SUBAPPLICATION SERVER_0_QO (* OPC-UA-Methode ohne Argumente (CREATE_METHOD): IND nur bei echtem Aufruf (QO=TRUE), RSP intern *)
  (* Standard: 61499-2; Description: Copyright (c) 2026 Meisterschulen am Ostbahnhof This program and the accompanying materials are made available under the terms of the Eclipse Public License 2.0 which is available at https://www.eclipse.org/legal/epl-2.0/ SPDX-License-Identifier: EPL-2.0 *)
  (* Version 1.0, 2026-11-25, Franz Höpfinger, Meisterschulen am Ostbahnhof, Neu: SERVER_0 + E_PERMIT(PERMIT=QO). Ein gescheitertes RSP meldet IND mit QO=FALSE, direkt IND->RSP ergab eine Endlosschleife. *)
  PACKAGE MyLib::net;
  (* Documentation:
  OPC-UA-Methode ohne Argumente, sicher beantwortet
   SERVER_0 mit CREATE_METHOD. IND geht nur bei QO = TRUE an RSP und nach außen (E_PERMIT).
   Warum: Findet FORTE zu einem RSP keinen offenen Aufruf (z. B. Antwort nach dem 4-s-Timeout), meldet der SERVER sofort wieder IND mit QO = FALSE. Direkt IND→RSP verdrahtet wird das eine Endlosschleife, die jede Runde die Aktion erneut auslöst (gesehen 2026-11-25, Boot-Zähler STG1).
   INIT darf unverbunden bleiben: SERVER.INIT ist selbst EInit, E_TRIG löst ihn im fboot aus.
  *)
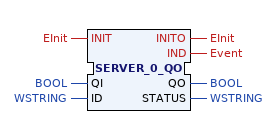
  EVENT_INPUT
    INIT : EInit; (* Initialization Request *)
  END_EVENT
  EVENT_OUTPUT
    INITO : EInit; (* Initialization Confirm *)
    IND; (* Methode wurde aufgerufen *)
  END_EVENT
  VAR_INPUT
    QI : BOOL := TRUE; (* Quality Input - TRUE to enable service *)
    ID : WSTRING; (* opc_ua[CREATE_METHOD;...] *)
  END_VAR
  VAR_OUTPUT
    QO : BOOL; (* Quality Output *)
    STATUS : WSTRING; (* Service Status *)
  END_VAR
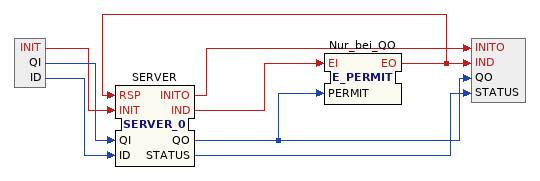
  FBS
    SERVER : iec61499::net::SERVER_0;
    Nur_bei_QO : iec61499::events::E_PERMIT; (* nur echter Call (QO=TRUE) *)
  END_FBS
  EVENT_CONNECTIONS
    SERVER.INITO TO INITO;
    SERVER.IND TO Nur_bei_QO.EI;
    Nur_bei_QO.EO TO SERVER.RSP;
    Nur_bei_QO.EO TO IND;
    INIT TO SERVER.INIT;
  END_CONNECTIONS
  DATA_CONNECTIONS
    QI TO SERVER.QI;
    ID TO SERVER.ID;
    SERVER.QO TO Nur_bei_QO.PERMIT;
    SERVER.QO TO QO;
    SERVER.STATUS TO STATUS;
  END_CONNECTIONS
END_SUBAPPLICATION
